TYPE "st_Io_Ph_DigitalInputs"
VERSION : 0.1
   STRUCT
      Zone1_K7k5Ss_Open { ExternalAccessible := 'False'; ExternalVisible := 'False'; ExternalWritable := 'False'; S7_SetPoint := 'False'} : "st_Io_Ph_DigitalInput";
      Zone1_K7k5Ss_Closed { ExternalAccessible := 'False'; ExternalVisible := 'False'; ExternalWritable := 'False'; S7_SetPoint := 'False'} : "st_Io_Ph_DigitalInput";
      Zone1_K7k5Vfd_Open { ExternalAccessible := 'False'; ExternalVisible := 'False'; ExternalWritable := 'False'; S7_SetPoint := 'False'} : "st_Io_Ph_DigitalInput";
      Zone1_K7k5Vfd_Closed { ExternalAccessible := 'False'; ExternalVisible := 'False'; ExternalWritable := 'False'; S7_SetPoint := 'False'} : "st_Io_Ph_DigitalInput";
      Zone1_K37Ss_Open { ExternalAccessible := 'False'; ExternalVisible := 'False'; ExternalWritable := 'False'; S7_SetPoint := 'False'} : "st_Io_Ph_DigitalInput";
      Zone1_K37Ss_Closed { ExternalAccessible := 'False'; ExternalVisible := 'False'; ExternalWritable := 'False'; S7_SetPoint := 'False'} : "st_Io_Ph_DigitalInput";
      Zone1_K37Vfd_Open { ExternalAccessible := 'False'; ExternalVisible := 'False'; ExternalWritable := 'False'; S7_SetPoint := 'False'} : "st_Io_Ph_DigitalInput";
      Zone1_K37Vfd_Closed { ExternalAccessible := 'False'; ExternalVisible := 'False'; ExternalWritable := 'False'; S7_SetPoint := 'False'} : "st_Io_Ph_DigitalInput";
      Zone1_K110Ss_Open { ExternalAccessible := 'False'; ExternalVisible := 'False'; ExternalWritable := 'False'; S7_SetPoint := 'False'} : "st_Io_Ph_DigitalInput";
      Zone1_K110Ss_Closed { ExternalAccessible := 'False'; ExternalVisible := 'False'; ExternalWritable := 'False'; S7_SetPoint := 'False'} : "st_Io_Ph_DigitalInput";
      Zone1_K110Vfd_Open { ExternalAccessible := 'False'; ExternalVisible := 'False'; ExternalWritable := 'False'; S7_SetPoint := 'False'} : "st_Io_Ph_DigitalInput";
      Zone1_K110Vfd_Closed { ExternalAccessible := 'False'; ExternalVisible := 'False'; ExternalWritable := 'False'; S7_SetPoint := 'False'} : "st_Io_Ph_DigitalInput";
      Zone1_Q560Ss_Open { ExternalAccessible := 'False'; ExternalVisible := 'False'; ExternalWritable := 'False'; S7_SetPoint := 'False'} : "st_Io_Ph_DigitalInput";
      Zone1_Q560Ss_Closed { ExternalAccessible := 'False'; ExternalVisible := 'False'; ExternalWritable := 'False'; S7_SetPoint := 'False'} : "st_Io_Ph_DigitalInput";
      Zone1_Q560Ss_SpringCharged { ExternalAccessible := 'False'; ExternalVisible := 'False'; ExternalWritable := 'False'; S7_SetPoint := 'False'} : "st_Io_Ph_DigitalInput";
      Zone1_Q630Vfd_Open { ExternalAccessible := 'False'; ExternalVisible := 'False'; ExternalWritable := 'False'; S7_SetPoint := 'False'} : "st_Io_Ph_DigitalInput";
      Zone1_Q630Vfd_Closed { ExternalAccessible := 'False'; ExternalVisible := 'False'; ExternalWritable := 'False'; S7_SetPoint := 'False'} : "st_Io_Ph_DigitalInput";
      Zone1_Q630Vfd_SpringCharged { ExternalAccessible := 'False'; ExternalVisible := 'False'; ExternalWritable := 'False'; S7_SetPoint := 'False'} : "st_Io_Ph_DigitalInput";
      Zone1_PendantStart { ExternalAccessible := 'False'; ExternalVisible := 'False'; ExternalWritable := 'False'; S7_SetPoint := 'False'} : "st_Io_Ph_DigitalInput";
      Zone1_PendantStop { ExternalAccessible := 'False'; ExternalVisible := 'False'; ExternalWritable := 'False'; S7_SetPoint := 'False'} : "st_Io_Ph_DigitalInput";
      Zone1_PendantTakeSample { ExternalAccessible := 'False'; ExternalVisible := 'False'; ExternalWritable := 'False'; S7_SetPoint := 'False'} : "st_Io_Ph_DigitalInput";
      Zone1_EStopOk { ExternalAccessible := 'False'; ExternalVisible := 'False'; ExternalWritable := 'False'; S7_SetPoint := 'False'} : "st_Io_Ph_DigitalInput";
      Zone1_PanelEStopOk { ExternalAccessible := 'False'; ExternalVisible := 'False'; ExternalWritable := 'False'; S7_SetPoint := 'False'} : "st_Io_Ph_DigitalInput";
      Zone2_K7k5Ss_Open { ExternalAccessible := 'False'; ExternalVisible := 'False'; ExternalWritable := 'False'; S7_SetPoint := 'False'} : "st_Io_Ph_DigitalInput";
      Zone2_K7k5Ss_Closed { ExternalAccessible := 'False'; ExternalVisible := 'False'; ExternalWritable := 'False'; S7_SetPoint := 'False'} : "st_Io_Ph_DigitalInput";
      Zone2_K7k5Vfd_Open { ExternalAccessible := 'False'; ExternalVisible := 'False'; ExternalWritable := 'False'; S7_SetPoint := 'False'} : "st_Io_Ph_DigitalInput";
      Zone2_K7k5Vfd_Closed { ExternalAccessible := 'False'; ExternalVisible := 'False'; ExternalWritable := 'False'; S7_SetPoint := 'False'} : "st_Io_Ph_DigitalInput";
      Zone2_K37Ss_Open { ExternalAccessible := 'False'; ExternalVisible := 'False'; ExternalWritable := 'False'; S7_SetPoint := 'False'} : "st_Io_Ph_DigitalInput";
      Zone2_K37Ss_Closed { ExternalAccessible := 'False'; ExternalVisible := 'False'; ExternalWritable := 'False'; S7_SetPoint := 'False'} : "st_Io_Ph_DigitalInput";
      Zone2_K37Vfd_Open { ExternalAccessible := 'False'; ExternalVisible := 'False'; ExternalWritable := 'False'; S7_SetPoint := 'False'} : "st_Io_Ph_DigitalInput";
      Zone2_K37Vfd_Closed { ExternalAccessible := 'False'; ExternalVisible := 'False'; ExternalWritable := 'False'; S7_SetPoint := 'False'} : "st_Io_Ph_DigitalInput";
      Zone2_K110Ss_Open { ExternalAccessible := 'False'; ExternalVisible := 'False'; ExternalWritable := 'False'; S7_SetPoint := 'False'} : "st_Io_Ph_DigitalInput";
      Zone2_K110Ss_Closed { ExternalAccessible := 'False'; ExternalVisible := 'False'; ExternalWritable := 'False'; S7_SetPoint := 'False'} : "st_Io_Ph_DigitalInput";
      Zone2_K110Vfd_Open { ExternalAccessible := 'False'; ExternalVisible := 'False'; ExternalWritable := 'False'; S7_SetPoint := 'False'} : "st_Io_Ph_DigitalInput";
      Zone2_K110Vfd_Closed { ExternalAccessible := 'False'; ExternalVisible := 'False'; ExternalWritable := 'False'; S7_SetPoint := 'False'} : "st_Io_Ph_DigitalInput";
      Zone2_Q560Ss_Open { ExternalAccessible := 'False'; ExternalVisible := 'False'; ExternalWritable := 'False'; S7_SetPoint := 'False'} : "st_Io_Ph_DigitalInput";
      Zone2_Q560Ss_Closed { ExternalAccessible := 'False'; ExternalVisible := 'False'; ExternalWritable := 'False'; S7_SetPoint := 'False'} : "st_Io_Ph_DigitalInput";
      Zone2_Q560Ss_SpringCharged { ExternalAccessible := 'False'; ExternalVisible := 'False'; ExternalWritable := 'False'; S7_SetPoint := 'False'} : "st_Io_Ph_DigitalInput";
      Zone2_Q630Vfd_Open { ExternalAccessible := 'False'; ExternalVisible := 'False'; ExternalWritable := 'False'; S7_SetPoint := 'False'} : "st_Io_Ph_DigitalInput";
      Zone2_Q630Vfd_Closed { ExternalAccessible := 'False'; ExternalVisible := 'False'; ExternalWritable := 'False'; S7_SetPoint := 'False'} : "st_Io_Ph_DigitalInput";
      Zone2_Q630Vfd_SpringCharged { ExternalAccessible := 'False'; ExternalVisible := 'False'; ExternalWritable := 'False'; S7_SetPoint := 'False'} : "st_Io_Ph_DigitalInput";
      Zone2_PendantStart { ExternalAccessible := 'False'; ExternalVisible := 'False'; ExternalWritable := 'False'; S7_SetPoint := 'False'} : "st_Io_Ph_DigitalInput";
      Zone2_PendantStop { ExternalAccessible := 'False'; ExternalVisible := 'False'; ExternalWritable := 'False'; S7_SetPoint := 'False'} : "st_Io_Ph_DigitalInput";
      Zone2_PendantTakeSample { ExternalAccessible := 'False'; ExternalVisible := 'False'; ExternalWritable := 'False'; S7_SetPoint := 'False'} : "st_Io_Ph_DigitalInput";
      Zone2_EStopOk { ExternalAccessible := 'False'; ExternalVisible := 'False'; ExternalWritable := 'False'; S7_SetPoint := 'False'} : "st_Io_Ph_DigitalInput";
      Zone2_PanelEStopOk { ExternalAccessible := 'False'; ExternalVisible := 'False'; ExternalWritable := 'False'; S7_SetPoint := 'False'} : "st_Io_Ph_DigitalInput";
      Zone3_K7k5Ss_Open { ExternalAccessible := 'False'; ExternalVisible := 'False'; ExternalWritable := 'False'; S7_SetPoint := 'False'} : "st_Io_Ph_DigitalInput";
      Zone3_K7k5Ss_Closed { ExternalAccessible := 'False'; ExternalVisible := 'False'; ExternalWritable := 'False'; S7_SetPoint := 'False'} : "st_Io_Ph_DigitalInput";
      Zone3_K7k5Vfd_Open { ExternalAccessible := 'False'; ExternalVisible := 'False'; ExternalWritable := 'False'; S7_SetPoint := 'False'} : "st_Io_Ph_DigitalInput";
      Zone3_K7k5Vfd_Closed { ExternalAccessible := 'False'; ExternalVisible := 'False'; ExternalWritable := 'False'; S7_SetPoint := 'False'} : "st_Io_Ph_DigitalInput";
      Zone3_K37Ss_Open { ExternalAccessible := 'False'; ExternalVisible := 'False'; ExternalWritable := 'False'; S7_SetPoint := 'False'} : "st_Io_Ph_DigitalInput";
      Zone3_K37Ss_Closed { ExternalAccessible := 'False'; ExternalVisible := 'False'; ExternalWritable := 'False'; S7_SetPoint := 'False'} : "st_Io_Ph_DigitalInput";
      Zone3_K37Vfd_Open { ExternalAccessible := 'False'; ExternalVisible := 'False'; ExternalWritable := 'False'; S7_SetPoint := 'False'} : "st_Io_Ph_DigitalInput";
      Zone3_K37Vfd_Closed { ExternalAccessible := 'False'; ExternalVisible := 'False'; ExternalWritable := 'False'; S7_SetPoint := 'False'} : "st_Io_Ph_DigitalInput";
      Zone3_K110Ss_Open { ExternalAccessible := 'False'; ExternalVisible := 'False'; ExternalWritable := 'False'; S7_SetPoint := 'False'} : "st_Io_Ph_DigitalInput";
      Zone3_K110Ss_Closed { ExternalAccessible := 'False'; ExternalVisible := 'False'; ExternalWritable := 'False'; S7_SetPoint := 'False'} : "st_Io_Ph_DigitalInput";
      Zone3_K110Vfd_Open { ExternalAccessible := 'False'; ExternalVisible := 'False'; ExternalWritable := 'False'; S7_SetPoint := 'False'} : "st_Io_Ph_DigitalInput";
      Zone3_K110Vfd_Closed { ExternalAccessible := 'False'; ExternalVisible := 'False'; ExternalWritable := 'False'; S7_SetPoint := 'False'} : "st_Io_Ph_DigitalInput";
      Zone3_Q560Ss_Open { ExternalAccessible := 'False'; ExternalVisible := 'False'; ExternalWritable := 'False'; S7_SetPoint := 'False'} : "st_Io_Ph_DigitalInput";
      Zone3_Q560Ss_Closed { ExternalAccessible := 'False'; ExternalVisible := 'False'; ExternalWritable := 'False'; S7_SetPoint := 'False'} : "st_Io_Ph_DigitalInput";
      Zone3_Q560Ss_SpringCharged { ExternalAccessible := 'False'; ExternalVisible := 'False'; ExternalWritable := 'False'; S7_SetPoint := 'False'} : "st_Io_Ph_DigitalInput";
      Zone3_Q630Vfd_Open { ExternalAccessible := 'False'; ExternalVisible := 'False'; ExternalWritable := 'False'; S7_SetPoint := 'False'} : "st_Io_Ph_DigitalInput";
      Zone3_Q630Vfd_Closed { ExternalAccessible := 'False'; ExternalVisible := 'False'; ExternalWritable := 'False'; S7_SetPoint := 'False'} : "st_Io_Ph_DigitalInput";
      Zone3_Q630Vfd_SpringCharged { ExternalAccessible := 'False'; ExternalVisible := 'False'; ExternalWritable := 'False'; S7_SetPoint := 'False'} : "st_Io_Ph_DigitalInput";
      Zone3_PendantStart { ExternalAccessible := 'False'; ExternalVisible := 'False'; ExternalWritable := 'False'; S7_SetPoint := 'False'} : "st_Io_Ph_DigitalInput";
      Zone3_PendantStop { ExternalAccessible := 'False'; ExternalVisible := 'False'; ExternalWritable := 'False'; S7_SetPoint := 'False'} : "st_Io_Ph_DigitalInput";
      Zone3_PendantTakeSample { ExternalAccessible := 'False'; ExternalVisible := 'False'; ExternalWritable := 'False'; S7_SetPoint := 'False'} : "st_Io_Ph_DigitalInput";
      Zone3_EStopOk { ExternalAccessible := 'False'; ExternalVisible := 'False'; ExternalWritable := 'False'; S7_SetPoint := 'False'} : "st_Io_Ph_DigitalInput";
      Zone3_PanelEStopOk { ExternalAccessible := 'False'; ExternalVisible := 'False'; ExternalWritable := 'False'; S7_SetPoint := 'False'} : "st_Io_Ph_DigitalInput";
      Drive_7k5Ss_Running { ExternalAccessible := 'False'; ExternalVisible := 'False'; ExternalWritable := 'False'; S7_SetPoint := 'False'} : "st_Io_Ph_DigitalInput";
      Drive_7k5Ss_Fault { ExternalAccessible := 'False'; ExternalVisible := 'False'; ExternalWritable := 'False'; S7_SetPoint := 'False'} : "st_Io_Ph_DigitalInput";
      Drive_7k5Vfd_Running { ExternalAccessible := 'False'; ExternalVisible := 'False'; ExternalWritable := 'False'; S7_SetPoint := 'False'} : "st_Io_Ph_DigitalInput";
      Drive_7k5Vfd_Fault { ExternalAccessible := 'False'; ExternalVisible := 'False'; ExternalWritable := 'False'; S7_SetPoint := 'False'} : "st_Io_Ph_DigitalInput";
      Drive_37Ss_Running { ExternalAccessible := 'False'; ExternalVisible := 'False'; ExternalWritable := 'False'; S7_SetPoint := 'False'} : "st_Io_Ph_DigitalInput";
      Drive_37Ss_Fault { ExternalAccessible := 'False'; ExternalVisible := 'False'; ExternalWritable := 'False'; S7_SetPoint := 'False'} : "st_Io_Ph_DigitalInput";
      Drive_37Vfd_Running { ExternalAccessible := 'False'; ExternalVisible := 'False'; ExternalWritable := 'False'; S7_SetPoint := 'False'} : "st_Io_Ph_DigitalInput";
      Drive_37Vfd_Fault { ExternalAccessible := 'False'; ExternalVisible := 'False'; ExternalWritable := 'False'; S7_SetPoint := 'False'} : "st_Io_Ph_DigitalInput";
      Drive_110Ss_Running { ExternalAccessible := 'False'; ExternalVisible := 'False'; ExternalWritable := 'False'; S7_SetPoint := 'False'} : "st_Io_Ph_DigitalInput";
      Drive_110Ss_Fault { ExternalAccessible := 'False'; ExternalVisible := 'False'; ExternalWritable := 'False'; S7_SetPoint := 'False'} : "st_Io_Ph_DigitalInput";
      Drive_110Vfd_Running { ExternalAccessible := 'False'; ExternalVisible := 'False'; ExternalWritable := 'False'; S7_SetPoint := 'False'} : "st_Io_Ph_DigitalInput";
      Drive_110Vfd_Fault { ExternalAccessible := 'False'; ExternalVisible := 'False'; ExternalWritable := 'False'; S7_SetPoint := 'False'} : "st_Io_Ph_DigitalInput";
      Drive_560Ss_Running { ExternalAccessible := 'False'; ExternalVisible := 'False'; ExternalWritable := 'False'; S7_SetPoint := 'False'} : "st_Io_Ph_DigitalInput";
      Drive_560Ss_Fault { ExternalAccessible := 'False'; ExternalVisible := 'False'; ExternalWritable := 'False'; S7_SetPoint := 'False'} : "st_Io_Ph_DigitalInput";
      Drive_630Vfd_Running { ExternalAccessible := 'False'; ExternalVisible := 'False'; ExternalWritable := 'False'; S7_SetPoint := 'False'} : "st_Io_Ph_DigitalInput";
      Drive_630Vfd_Fault { ExternalAccessible := 'False'; ExternalVisible := 'False'; ExternalWritable := 'False'; S7_SetPoint := 'False'} : "st_Io_Ph_DigitalInput";
   END_STRUCT;

END_TYPE

